Staubli VAL3: _bindPROG.pgx

program _bindPROG(string x_sHtml)
  local num l_i
  local string l_sbtn
begin
  for l_i = 1 to 6
    l_sbtn="btn"+toString("",l_i)
    userPageBindClick(x_sHtml,l_sbtn,bInsert[l_i],true)
  endFor

  userPageBind(x_sHtml,"lbl1","innerHTML",sPgIndexPROG,1,"r")
  userPageBind(x_sHtml,"lbl2","innerHTML",sPagePROG,1,"r")

  userPageBindClick(x_sHtml,"btn7",bSelProg,true)
  userPageBindClick(x_sHtml,"btn8",bSelTraj,true)
  userPageBind(x_sHtml,"lst1","value",sInsertItem,1,"rw")

end
